Fanuc KAREL source: kt00408.KL

-- PROVISIONAL review KL for V1013-1; original PC SHA256 bf0c4b1b3bf633a90c65d32cc1ea66bb213b93fdb27c0a926f7662ce418c76a0
-- Incomplete behavior may be omitted. Consult companion uncertainty JSON. Do not deploy.
PROGRAM KT00408
%NOLOCKGROUP
VAR
  R1 : REAL
  OUT : BOOLEAN
-- UNRESOLVED_DECL H2 type=002017
BEGIN
  -- UNRESOLVED_PC offsets 5-16; opcodes 2E,23
  -- UNRESOLVED_PC offsets 21-35; opcodes 2E,22,9D,33,B4
  -- UNRESOLVED_PC offsets 40-63; opcodes 21,22,9D,33,B3,64,71,23
  -- UNRESOLVED_PC offsets 68-72; opcodes 7F
END KT00408
